(* IEC 61131-3 sources: codesys-framework/txt/application/WeVe Core (library)/60 Event/FB_Event, 3 files *)

(* ---- Condition.method.st ---- *)
// Elke cyclus aanroepen voor een warning of alarm.
//   stijgende flank : event wordt actief en logt 'raised' (met scPayload)
//   dalende flank   : logt 'cleared'
//                     niet resetbaar -> event wordt meteen inactief
//                     resetbaar      -> event blijft actief tot Reset()
// Geeft Active terug.
METHOD Condition : BOOL
VAR_INPUT
	xCondition 		: BOOL;
	scPayload 		: SC_EventPayload := (asPayload := [10('')]);	// mag weggelaten worden
END_VAR

// --- BEGIN IMPLEMENTATION ---

IF _xDisabled THEN
	Condition := FALSE;
	RETURN;
END_IF

// Stijgende flank
IF xCondition AND NOT _xCondition THEN
	_xActive := TRUE;
	_scPayload := scPayload;
	WriteLog(sTransition := 'raised', scPayload := _scPayload);

// Dalende flank
ELSIF NOT xCondition AND _xCondition THEN
	WriteLog(sTransition := 'cleared', scPayload := _scPayload);

	IF NOT _scConfig.xResetable THEN
		_xActive := FALSE;
	END_IF

END_IF

_xCondition := xCondition;
Condition := _xActive;

(* ---- Log.method.st ---- *)
// Eenmalige melding, bv. drukknop of aanvraag. Houdt geen toestand bij.
// TRUE = gelogd. FALSE = uitgeschakeld, geen logger of buffer vol.
METHOD Log : BOOL
VAR_INPUT
	scPayload 		: SC_EventPayload := (asPayload := [10('')]);	// mag weggelaten worden
END_VAR

// --- BEGIN IMPLEMENTATION ---

IF _xDisabled THEN
	Log := FALSE;
	RETURN;
END_IF

Log := WriteLog(sTransition := '', scPayload := scPayload);

(* ---- Reset.method.st ---- *)
// Reset het event, maar enkel als de conditie weg is. Logt 'reset'.
// TRUE = event is niet (meer) actief.
METHOD Reset : BOOL
VAR_INPUT
END_VAR

// --- BEGIN IMPLEMENTATION ---

IF NOT _xActive THEN
	Reset := TRUE;
	RETURN;
END_IF

// Oorzaak nog aanwezig: reset weigeren
IF _xCondition THEN
	Reset := FALSE;
	RETURN;
END_IF

_xActive := FALSE;
WriteLog(sTransition := 'reset', scPayload := _scPayload);
Reset := TRUE;
